RoboDK station: PickPlace_Delta_ABB.rdk

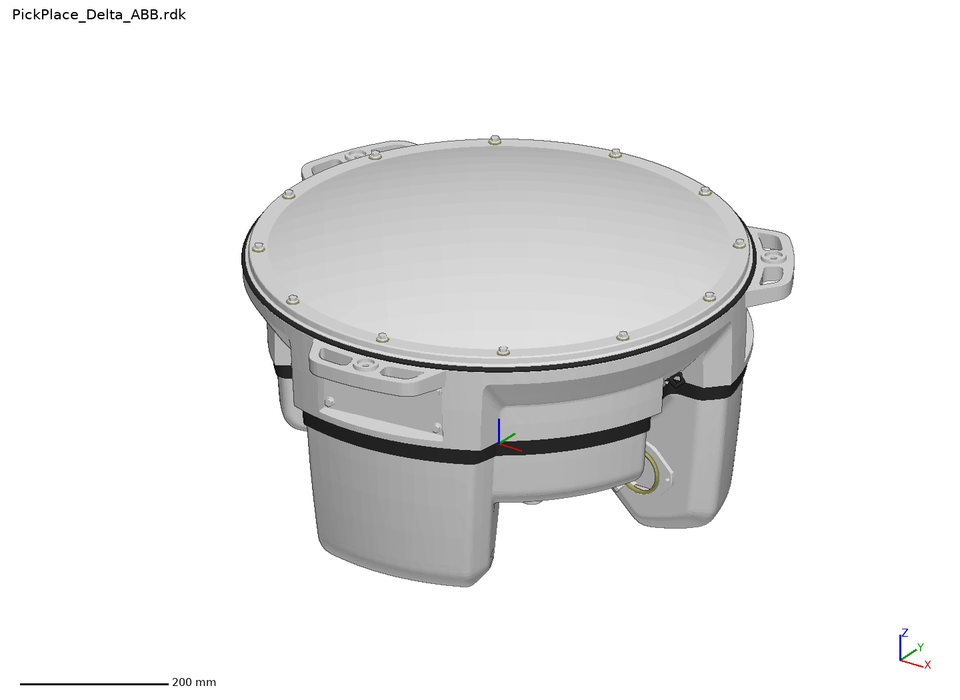
[picture v0: the station drawn from its stored meshes, robots at their saved joint values, targets as dots, program paths as lines]
Station PickPlace_Delta_ABB (saved by RoboDK 6.0.1). Poses are relative to the parent item; angles as X-Y-Z fixed-axis rotations.
Station parameters (name, value as stored): SICK WL4S Laser Sensor, 0, start_prox, 0
  - frame Conveyor Belt Wide (2m) Base at (0, 0, -10) mm
    - robot Conveyor Belt Wide (2m): 1 axes
        modified DH rows (alpha deg, a mm, theta deg, d mm): 0, 0, 0, 0 linear
        base shift (0, 0, 0) mm, rotated rx 0 ry 90 rz 0 deg
        joint limits [-900000] to [900000]; home [0]; saved at [-824508]
      - frame Conveyor Frame at (1954.3, 0, -10) mm
        - object Box at (897730.69, 156.17, 12.65) mm, rotated rx -0.59 ry -0.06 rz -23.58 deg, size 10 x 20 x 5 mm, geometry from box.sld
        - object Box at (897637.69, 177.81, 12.44) mm, rotated rx -0.3 ry 0.51 rz 41.51 deg, size 10 x 20 x 5 mm, geometry from box.sld
        - object Box at (897468.69, 142.01, 12.79) mm, rotated rx -0.52 ry 0.28 rz 10.42 deg, size 10 x 20 x 5 mm, geometry from box.sld
        - object Box at (897370.7, 94.71, 13.25) mm, rotated rx -0.59 ry 0.03 rz -15.02 deg, size 10 x 20 x 5 mm, geometry from box.sld
        - object Box at (897268.7, 59.56, 13.6) mm, rotated rx -0.59 ry -0.09 rz -26.61 deg, size 10 x 20 x 5 mm, geometry from box.sld
        - object Box at (897066.69, 179.61, 12.42) mm, rotated rx -0.4 ry 0.44 rz 29.48 deg, size 10 x 20 x 5 mm, geometry from box.sld
        - object Box at (896960.69, 179.12, 12.42) mm, rotated rx -0.29 ry 0.52 rz 42.93 deg, size 10 x 20 x 5 mm, geometry from box.sld
        - object Box at (896886.7, 104.97, 13.15) mm, rotated rx -0.55 ry 0.22 rz 3.61 deg, size 10 x 20 x 5 mm, geometry from box.sld
        - object Box at (896794.7, 36.7, 13.82) mm, rotated rx -0.43 ry 0.41 rz 25.81 deg, size 10 x 20 x 5 mm, geometry from box.sld
        - object Box at (896686.7, 102.36, 13.18) mm, rotated rx -0.56 ry -0.21 rz -38.82 deg, size 10 x 20 x 5 mm, geometry from box.sld
        - object Box at (896480.69, 181.98, 12.39) mm, rotated rx -0.53 ry -0.26 rz -44.04 deg, size 10 x 20 x 5 mm, geometry from box.sld
        - object Box at (896386.7, 69.3, 13.5) mm, rotated rx -0.54 ry -0.24 rz -42.5 deg, size 10 x 20 x 5 mm, geometry from box.sld
        - object Box at (896271.7, 21, 13.98) mm, rotated rx -0.57 ry -0.15 rz -32.81 deg, size 10 x 20 x 5 mm, geometry from box.sld
        - object Box at (896066.7, 121.17, 12.99) mm, rotated rx -0.58 ry 0.12 rz -6.35 deg, size 10 x 20 x 5 mm, geometry from box.sld
        - object Box at (895875.7, 101.57, 13.19) mm, rotated rx -0.59 ry -0.02 rz -20.07 deg, size 10 x 20 x 5 mm, geometry from box.sld
        - object Box at (895769.69, 140.05, 12.81) mm, rotated rx -0.59 ry 0.01 rz -17.18 deg, size 10 x 20 x 5 mm, geometry from box.sld
        - object Box at (895559.7, 47.66, 13.72) mm, rotated rx -0.46 ry 0.38 rz 21.06 deg, size 10 x 20 x 5 mm, geometry from box.sld
        - object Box at (895483.69, 179.87, 12.41) mm, rotated rx -0.56 ry 0.2 rz 1.63 deg, size 10 x 20 x 5 mm, geometry from box.sld
        - object Box at (895370.7, 123.7, 12.97) mm, rotated rx -0.59 ry 0.04 rz -14.74 deg, size 10 x 20 x 5 mm, geometry from box.sld
        - object Box at (895264.7, 131.8, 12.89) mm, rotated rx -0.58 ry -0.14 rz -31.52 deg, size 10 x 20 x 5 mm, geometry from box.sld
        - object Box at (895176.7, 127.41, 12.93) mm, rotated rx -0.59 ry -0.01 rz -19.42 deg, size 10 x 20 x 5 mm, geometry from box.sld
        - object Box at (895070.69, 148.83, 12.72) mm, rotated rx -0.59 ry 0.04 rz -13.82 deg, size 10 x 20 x 5 mm, geometry from box.sld
        - object Box at (894830.7, 134.47, 12.86) mm, rotated rx -0.55 ry -0.21 rz -39.3 deg, size 10 x 20 x 5 mm, geometry from box.sld
        - object Box at (894736.69, 145.17, 12.76) mm, rotated rx -0.58 ry 0.12 rz -6.93 deg, size 10 x 20 x 5 mm, geometry from box.sld
        - object Box at (894651.7, 66.02, 13.54) mm, rotated rx -0.57 ry -0.15 rz -32.83 deg, size 10 x 20 x 5 mm, geometry from box.sld
        - object Box at (894556.7, 45.28, 13.74) mm, rotated rx -0.42 ry 0.42 rz 26.95 deg, size 10 x 20 x 5 mm, geometry from box.sld
        - object Box at (894429.7, 71.11, 13.49) mm, rotated rx -0.56 ry -0.2 rz -37.64 deg, size 10 x 20 x 5 mm, geometry from box.sld
        - object Box at (894341.69, 182.71, 12.39) mm, rotated rx -0.59 ry 0.01 rz -17.44 deg, size 10 x 20 x 5 mm, geometry from box.sld
        - object Box at (894244.7, 91.87, 13.28) mm, rotated rx -0.54 ry -0.24 rz -42.33 deg, size 10 x 20 x 5 mm, geometry from box.sld
        - object Box at (893942.7, 111.28, 13.09) mm, rotated rx -0.52 ry 0.28 rz 9.97 deg, size 10 x 20 x 5 mm, geometry from box.sld
        - object Box at (893859.7, 78.43, 13.41) mm, rotated rx -0.59 ry 0.05 rz -12.95 deg, size 10 x 20 x 5 mm, geometry from box.sld
        - object Box at (893731.69, 182.25, 12.39) mm, rotated rx -0.59 ry -0.05 rz -23.07 deg, size 10 x 20 x 5 mm, geometry from box.sld
        - object Box at (893626.69, 198.26, 12.23) mm, rotated rx -0.44 ry 0.4 rz 24.46 deg, size 10 x 20 x 5 mm, geometry from box.sld
        - object Box at (893339.7, 130.91, 12.9) mm, rotated rx -0.43 ry 0.41 rz 25.41 deg, size 10 x 20 x 5 mm, geometry from box.sld
        - object Box at (893114.69, 144.51, 12.76) mm, rotated rx -0.59 ry -0.04 rz -22.45 deg, size 10 x 20 x 5 mm, geometry from box.sld
        - object Box at (893046.7, 53.65, 13.66) mm, rotated rx -0.57 ry 0.15 rz -3.55 deg, size 10 x 20 x 5 mm, geometry from box.sld
        - object Box at (892837.69, 193.79, 12.28) mm, rotated rx -0.41 ry 0.43 rz 28.71 deg, size 10 x 20 x 5 mm, geometry from box.sld
        - object Box at (892611.7, 108.11, 13.12) mm, rotated rx -0.42 ry 0.42 rz 26.96 deg, size 10 x 20 x 5 mm, geometry from box.sld
        - object Box at (892480.7, 68.86, 13.51) mm, rotated rx -0.51 ry 0.3 rz 12.73 deg, size 10 x 20 x 5 mm, geometry from box.sld
        - object Box at (892369.7, 112.85, 13.07) mm, rotated rx -0.59 ry 0.02 rz -16.52 deg, size 10 x 20 x 5 mm, geometry from box.sld
        - object Box at (892237.7, 18.64, 14) mm, rotated rx -0.59 ry 0.06 rz -11.95 deg, size 10 x 20 x 5 mm, geometry from box.sld
        - object Box at (892122.69, 158.92, 12.62) mm, rotated rx -0.43 ry 0.41 rz 25.04 deg, size 10 x 20 x 5 mm, geometry from box.sld
        - object Box at (892026.7, 94.47, 13.26) mm, rotated rx -0.59 ry 0.07 rz -11.43 deg, size 10 x 20 x 5 mm, geometry from box.sld
        - object Box at (891747.7, 66.89, 13.53) mm, rotated rx -0.59 ry -0.02 rz -20.16 deg, size 10 x 20 x 5 mm, geometry from box.sld
        - object Box at (891542.69, 140.71, 12.8) mm, rotated rx -0.42 ry 0.42 rz 26.92 deg, size 10 x 20 x 5 mm, geometry from box.sld
        - object Box at (891444.69, 197.73, 12.24) mm, rotated rx -0.3 ry 0.51 rz 41.43 deg, size 10 x 20 x 5 mm, geometry from box.sld
        - object Box at (891351.7, 42.87, 13.76) mm, rotated rx -0.54 ry -0.24 rz -41.92 deg, size 10 x 20 x 5 mm, geometry from box.sld
        - object Box at (891043.69, 177.02, 12.44) mm, rotated rx -0.57 ry -0.17 rz -35.25 deg, size 10 x 20 x 5 mm, geometry from box.sld
        - object Box at (890826.69, 146.16, 12.75) mm, rotated rx -0.57 ry -0.16 rz -33.48 deg, size 10 x 20 x 5 mm, geometry from box.sld
        - object Box at (890637.7, 55.66, 13.64) mm, rotated rx -0.58 ry -0.13 rz -30.72 deg, size 10 x 20 x 5 mm, geometry from box.sld
        - object Box at (890524.69, 170.49, 12.51) mm, rotated rx -0.57 ry -0.16 rz -33.37 deg, size 10 x 20 x 5 mm, geometry from box.sld
        - object Box at (890376.69, 167.1, 12.54) mm, rotated rx -0.58 ry -0.12 rz -30.29 deg, size 10 x 20 x 5 mm, geometry from box.sld
        - object Box at (890243.7, 28.37, 13.91) mm, rotated rx -0.59 ry -0.03 rz -21.44 deg, size 10 x 20 x 5 mm, geometry from box.sld
        - object Box at (890087.7, 32.55, 13.87) mm, rotated rx -0.58 ry -0.14 rz -31.77 deg, size 10 x 20 x 5 mm, geometry from box.sld
        - object Box at (889842.7, 52.41, 13.67) mm, rotated rx -0.49 ry 0.33 rz 15.68 deg, size 10 x 20 x 5 mm, geometry from box.sld
        - object Box at (889568.7, 81.43, 13.38) mm, rotated rx -0.43 ry 0.41 rz 25.3 deg, size 10 x 20 x 5 mm, geometry from box.sld
        - object Box at (889310.7, 27.98, 13.91) mm, rotated rx -0.57 ry 0.18 rz -0.36 deg, size 10 x 20 x 5 mm, geometry from box.sld
        - object Box at (889224.69, 159.39, 12.62) mm, rotated rx -0.5 ry 0.32 rz 14.94 deg, size 10 x 20 x 5 mm, geometry from box.sld
        - object Box at (888940.7, 109.26, 13.11) mm, rotated rx -0.58 ry 0.13 rz -5.05 deg, size 10 x 20 x 5 mm, geometry from box.sld
        - object Box at (888797.7, 63.43, 13.56) mm, rotated rx -0.32 ry 0.5 rz 38.96 deg, size 10 x 20 x 5 mm, geometry from box.sld
        - object Box at (888564.7, 67.11, 13.52) mm, rotated rx -0.39 ry 0.45 rz 31 deg, size 10 x 20 x 5 mm, geometry from box.sld
        - object Box at (888277.69, 157.91, 12.63) mm, rotated rx -0.51 ry 0.31 rz 12.91 deg, size 10 x 20 x 5 mm, geometry from box.sld
        - object Box at (888179.7, 88.13, 13.32) mm, rotated rx -0.53 ry 0.26 rz 8.19 deg, size 10 x 20 x 5 mm, geometry from box.sld
        - object Box at (888049.69, 160.71, 12.6) mm, rotated rx -0.59 ry -0.04 rz -22.46 deg, size 10 x 20 x 5 mm, geometry from box.sld
        - object Box at (887779.69, 175.73, 12.46) mm, rotated rx -0.56 ry 0.18 rz -0.25 deg, size 10 x 20 x 5 mm, geometry from box.sld
        - object Box at (887507.7, 34.78, 13.84) mm, rotated rx -0.55 ry 0.23 rz 5.02 deg, size 10 x 20 x 5 mm, geometry from box.sld
        - object Box at (887341.69, 183.19, 12.38) mm, rotated rx -0.35 ry 0.48 rz 36.16 deg, size 10 x 20 x 5 mm, geometry from box.sld
        - object Box at (887031.7, 18.9, 14) mm, rotated rx -0.59 ry -0.08 rz -26.28 deg, size 10 x 20 x 5 mm, geometry from box.sld
        - object Box at (886865.69, 175.99, 12.45) mm, rotated rx -0.58 ry 0.15 rz -3.88 deg, size 10 x 20 x 5 mm, geometry from box.sld
        - object Box at (886728.7, 132.72, 12.88) mm, rotated rx -0.47 ry 0.36 rz 18.81 deg, size 10 x 20 x 5 mm, geometry from box.sld
        - object Box at (886614.7, 70.74, 13.49) mm, rotated rx -0.56 ry 0.2 rz 1.77 deg, size 10 x 20 x 5 mm, geometry from box.sld
        - object Box at (886478.7, 44.32, 13.75) mm, rotated rx -0.58 ry -0.11 rz -29.31 deg, size 10 x 20 x 5 mm, geometry from box.sld
        - object Box at (886356.7, 71.95, 13.48) mm, rotated rx -0.51 ry 0.31 rz 13.14 deg, size 10 x 20 x 5 mm, geometry from box.sld
        - object Box at (886087.7, 108.74, 13.12) mm, rotated rx -0.58 ry -0.13 rz -31.01 deg, size 10 x 20 x 5 mm, geometry from box.sld
        - object Box at (885692.69, 167.79, 12.53) mm, rotated rx -0.59 ry -0.01 rz -18.94 deg, size 10 x 20 x 5 mm, geometry from box.sld
        - object Box at (885279.7, 93.51, 13.26) mm, rotated rx -0.57 ry -0.17 rz -35.18 deg, size 10 x 20 x 5 mm, geometry from box.sld
        - object Box at (885168.7, 33.77, 13.85) mm, rotated rx -0.59 ry 0.09 rz -9.53 deg, size 10 x 20 x 5 mm, geometry from box.sld
        - object Box at (884865.7, 95.2, 13.25) mm, rotated rx -0.59 ry -0.1 rz -27.76 deg, size 10 x 20 x 5 mm, geometry from box.sld
        - object Box at (884481.69, 195.64, 12.26) mm, rotated rx -0.59 ry 0.05 rz -13.6 deg, size 10 x 20 x 5 mm, geometry from box.sld
        - object Box at (884238.7, 13.58, 14.05) mm, rotated rx -0.29 ry 0.52 rz 42.46 deg, size 10 x 20 x 5 mm, geometry from box.sld
        - object Box at (883600.69, 168.73, 12.52) mm, rotated rx -0.39 ry 0.45 rz 31.19 deg, size 10 x 20 x 5 mm, geometry from box.sld
        - object Box at (883471.69, 175.1, 12.46) mm, rotated rx -0.56 ry -0.19 rz -36.67 deg, size 10 x 20 x 5 mm, geometry from box.sld
        - object Box at (883117.7, 8.08, 14.11) mm, rotated rx -0.59 ry 0 rz -18.33 deg, size 10 x 20 x 5 mm, geometry from box.sld
        - object Box at (882411.69, 148.37, 12.72) mm, rotated rx -0.37 ry 0.47 rz 33.68 deg, size 10 x 20 x 5 mm, geometry from box.sld
        - object Box at (881994.69, 149.13, 12.72) mm, rotated rx -0.55 ry -0.21 rz -39.37 deg, size 10 x 20 x 5 mm, geometry from box.sld
        - object Box at (881721.7, 36.8, 13.82) mm, rotated rx -0.56 ry -0.18 rz -36.26 deg, size 10 x 20 x 5 mm, geometry from box.sld
        - object Box at (881386.69, 181.59, 12.4) mm, rotated rx -0.48 ry 0.34 rz 17.23 deg, size 10 x 20 x 5 mm, geometry from box.sld
        - object Box at (881076.7, 104.94, 13.15) mm, rotated rx -0.58 ry 0.14 rz -4.54 deg, size 10 x 20 x 5 mm, geometry from box.sld
        - object Box at (880927.7, 105.79, 13.14) mm, rotated rx -0.59 ry -0.05 rz -23.21 deg, size 10 x 20 x 5 mm, geometry from box.sld
        - object Box at (880633.7, 82.69, 13.37) mm, rotated rx -0.58 ry 0.15 rz -3.91 deg, size 10 x 20 x 5 mm, geometry from box.sld
        - object Box at (880250.7, 100.17, 13.2) mm, rotated rx -0.35 ry 0.48 rz 36.02 deg, size 10 x 20 x 5 mm, geometry from box.sld
        - object Box at (879967.7, 8.92, 14.1) mm, rotated rx -0.34 ry 0.49 rz 36.88 deg, size 10 x 20 x 5 mm, geometry from box.sld
        - object Box at (879702.69, 197.41, 12.24) mm, rotated rx -0.54 ry 0.24 rz 5.94 deg, size 10 x 20 x 5 mm, geometry from box.sld
        - object Box at (879327.7, 134.52, 12.86) mm, rotated rx -0.31 ry 0.51 rz 40.25 deg, size 10 x 20 x 5 mm, geometry from box.sld
        - object Box at (879021.7, 66.06, 13.54) mm, rotated rx -0.59 ry -0.09 rz -26.74 deg, size 10 x 20 x 5 mm, geometry from box.sld
        - object Box at (878707.7, 123.22, 12.97) mm, rotated rx -0.3 ry 0.51 rz 41.76 deg, size 10 x 20 x 5 mm, geometry from box.sld
        - object Box at (878458.7, 26.6, 13.92) mm, rotated rx -0.38 ry 0.46 rz 32.24 deg, size 10 x 20 x 5 mm, geometry from box.sld
        - object Box at (878137.69, 148.25, 12.73) mm, rotated rx -0.36 ry 0.47 rz 34.26 deg, size 10 x 20 x 5 mm, geometry from box.sld
        - object Box at (877571.7, 84.32, 13.36) mm, rotated rx -0.33 ry 0.5 rz 38.45 deg, size 10 x 20 x 5 mm, geometry from box.sld
        - object Box at (877259.69, 194, 12.28) mm, rotated rx -0.49 ry 0.33 rz 15.69 deg, size 10 x 20 x 5 mm, geometry from box.sld
        - object Box at (877049.69, 140.02, 12.81) mm, rotated rx -0.59 ry 0.01 rz -17.21 deg, size 10 x 20 x 5 mm, geometry from box.sld
        - object Box at (876618.69, 160.9, 12.6) mm, rotated rx -0.56 ry -0.21 rz -38.5 deg, size 10 x 20 x 5 mm, geometry from box.sld
        - object Box at (876232.69, 160.62, 12.6) mm, rotated rx -0.52 ry 0.28 rz 10.27 deg, size 10 x 20 x 5 mm, geometry from box.sld
        - object Box at (876057.7, 87.66, 13.32) mm, rotated rx -0.56 ry -0.21 rz -38.4 deg, size 10 x 20 x 5 mm, geometry from box.sld
        - object Box at (875735.69, 153.67, 12.67) mm, rotated rx -0.57 ry 0.17 rz -1.28 deg, size 10 x 20 x 5 mm, geometry from box.sld
        - object Box at (875385.7, 12.69, 14.06) mm, rotated rx -0.52 ry 0.29 rz 10.64 deg, size 10 x 20 x 5 mm, geometry from box.sld
        - object Box at (874877.7, 46, 13.73) mm, rotated rx -0.46 ry 0.37 rz 20.28 deg, size 10 x 20 x 5 mm, geometry from box.sld
        - object Box at (874555.69, 151.65, 12.69) mm, rotated rx -0.58 ry -0.14 rz -31.99 deg, size 10 x 20 x 5 mm, geometry from box.sld
        - object Box at (873807.69, 173.16, 12.48) mm, rotated rx -0.28 ry 0.52 rz 43.49 deg, size 10 x 20 x 5 mm, geometry from box.sld
        - object Box at (872936.7, 49.92, 13.69) mm, rotated rx -0.34 ry 0.49 rz 36.91 deg, size 10 x 20 x 5 mm, geometry from box.sld
        - object Box at (872785.69, 161.75, 12.59) mm, rotated rx -0.59 ry 0.09 rz -9.24 deg, size 10 x 20 x 5 mm, geometry from box.sld
        - object Box at (872664.7, 91.07, 13.29) mm, rotated rx -0.52 ry 0.29 rz 11.2 deg, size 10 x 20 x 5 mm, geometry from box.sld
        - object Box at (872500.7, 40.63, 13.79) mm, rotated rx -0.59 ry 0.06 rz -12.41 deg, size 10 x 20 x 5 mm, geometry from box.sld
        - object Box at (872142.7, 105.29, 13.15) mm, rotated rx -0.5 ry 0.32 rz 14.54 deg, size 10 x 20 x 5 mm, geometry from box.sld
        - object Box at (871888.7, 15.8, 14.03) mm, rotated rx -0.53 ry -0.27 rz -44.74 deg, size 10 x 20 x 5 mm, geometry from box.sld
        - object Box at (871587.7, 7.86, 14.11) mm, rotated rx -0.51 ry 0.3 rz 12.38 deg, size 10 x 20 x 5 mm, geometry from box.sld
        - object Box at (870973.69, 136.14, 12.85) mm, rotated rx -0.42 ry 0.42 rz 26.47 deg, size 10 x 20 x 5 mm, geometry from box.sld
        - object Box at (869775.7, 70.75, 13.49) mm, rotated rx -0.38 ry 0.46 rz 32.57 deg, size 10 x 20 x 5 mm, geometry from box.sld
        - object Box at (869038.69, 182.24, 12.39) mm, rotated rx -0.55 ry -0.21 rz -39.23 deg, size 10 x 20 x 5 mm, geometry from box.sld
        - object Box at (868878.7, 50.82, 13.69) mm, rotated rx -0.59 ry 0.03 rz -15.61 deg, size 10 x 20 x 5 mm, geometry from box.sld
        - object Box at (868388.7, 14.54, 14.04) mm, rotated rx -0.57 ry 0.15 rz -3.36 deg, size 10 x 20 x 5 mm, geometry from box.sld
        - object Box at (867960.7, 83.04, 13.37) mm, rotated rx -0.52 ry 0.28 rz 9.96 deg, size 10 x 20 x 5 mm, geometry from box.sld
        - object Box at (867636.7, 10.32, 14.08) mm, rotated rx -0.4 ry 0.44 rz 29.65 deg, size 10 x 20 x 5 mm, geometry from box.sld
        - object Box at (867059.69, 162.68, 12.58) mm, rotated rx -0.58 ry -0.11 rz -28.52 deg, size 10 x 20 x 5 mm, geometry from box.sld
        - object Box at (866931.7, 128.82, 12.92) mm, rotated rx -0.55 ry 0.21 rz 2.62 deg, size 10 x 20 x 5 mm, geometry from box.sld
        - object Box at (866587.69, 156.78, 12.64) mm, rotated rx -0.47 ry 0.36 rz 19.55 deg, size 10 x 20 x 5 mm, geometry from box.sld
        - object Box at (866076.69, 184.18, 12.37) mm, rotated rx -0.59 ry 0.04 rz -14.44 deg, size 10 x 20 x 5 mm, geometry from box.sld
        - object Box at (865379.7, 5.34, 14.13) mm, rotated rx -0.58 ry -0.13 rz -30.77 deg, size 10 x 20 x 5 mm, geometry from box.sld
        - object Box at (865212.69, 149.76, 12.71) mm, rotated rx -0.56 ry -0.2 rz -38.32 deg, size 10 x 20 x 5 mm, geometry from box.sld
        - object Box at (864790.7, 7.34, 14.11) mm, rotated rx -0.59 ry 0.07 rz -11.85 deg, size 10 x 20 x 5 mm, geometry from box.sld
        - object Box at (864117.7, 14.14, 14.05) mm, rotated rx -0.4 ry 0.44 rz 29.12 deg, size 10 x 20 x 5 mm, geometry from box.sld
        - object Box at (864010.69, 143.76, 12.77) mm, rotated rx -0.59 ry 0 rz -18.52 deg, size 10 x 20 x 5 mm, geometry from box.sld
        - object Box at (863847.69, 186.35, 12.35) mm, rotated rx -0.54 ry -0.24 rz -42.33 deg, size 10 x 20 x 5 mm, geometry from box.sld
        - object Box at (863773.7, 56.85, 13.63) mm, rotated rx -0.53 ry -0.27 rz -44.81 deg, size 10 x 20 x 5 mm, geometry from box.sld
        - object Box at (863691.7, 42.47, 13.77) mm, rotated rx -0.57 ry -0.16 rz -34.11 deg, size 10 x 20 x 5 mm, geometry from box.sld
        - object Box at (863609.7, 44.95, 13.74) mm, rotated rx -0.5 ry 0.33 rz 15.05 deg, size 10 x 20 x 5 mm, geometry from box.sld
        - object Box at (863543.7, 34.25, 13.85) mm, rotated rx -0.51 ry 0.31 rz 13.03 deg, size 10 x 20 x 5 mm, geometry from box.sld
        - object Box at (863468.7, 76.02, 13.44) mm, rotated rx -0.59 ry 0.1 rz -8.77 deg, size 10 x 20 x 5 mm, geometry from box.sld
        - object Box at (863299.7, 107.42, 13.13) mm, rotated rx -0.55 ry -0.21 rz -39.28 deg, size 10 x 20 x 5 mm, geometry from box.sld
        - object Box at (863239.69, 195.88, 12.26) mm, rotated rx -0.29 ry 0.52 rz 42.8 deg, size 10 x 20 x 5 mm, geometry from box.sld
        - object Box at (863168.7, 58.58, 13.61) mm, rotated rx -0.58 ry 0.15 rz -3.89 deg, size 10 x 20 x 5 mm, geometry from box.sld
        - object Box at (863074.69, 157.27, 12.64) mm, rotated rx -0.57 ry 0.17 rz -1.09 deg, size 10 x 20 x 5 mm, geometry from box.sld
        - object Box at (862995.7, 21.42, 13.97) mm, rotated rx -0.59 ry 0.1 rz -8.62 deg, size 10 x 20 x 5 mm, geometry from box.sld
        - object Box at (862844.69, 190.46, 12.31) mm, rotated rx -0.47 ry 0.37 rz 19.8 deg, size 10 x 20 x 5 mm, geometry from box.sld
        - object Box at (862697.7, 12.52, 14.06) mm, rotated rx -0.55 ry 0.22 rz 3.49 deg, size 10 x 20 x 5 mm, geometry from box.sld
        - object Box at (862605.7, 93.15, 13.27) mm, rotated rx -0.43 ry 0.41 rz 25.14 deg, size 10 x 20 x 5 mm, geometry from box.sld
        - object Box at (862511.69, 173.93, 12.47) mm, rotated rx -0.49 ry 0.33 rz 15.38 deg, size 10 x 20 x 5 mm, geometry from box.sld
        - object Box at (862445.69, 170.13, 12.51) mm, rotated rx -0.56 ry -0.21 rz -38.76 deg, size 10 x 20 x 5 mm, geometry from box.sld
        - object Box at (862285.69, 194.2, 12.27) mm, rotated rx -0.59 ry -0.02 rz -20.35 deg, size 10 x 20 x 5 mm, geometry from box.sld
        - object Box at (862212.7, 48.11, 13.71) mm, rotated rx -0.53 ry 0.26 rz 8.23 deg, size 10 x 20 x 5 mm, geometry from box.sld
        - object Box at (862077.7, 40.74, 13.78) mm, rotated rx -0.57 ry -0.15 rz -33.02 deg, size 10 x 20 x 5 mm, geometry from box.sld
        - object Box at (862001.69, 144.78, 12.76) mm, rotated rx -0.59 ry -0.04 rz -21.98 deg, size 10 x 20 x 5 mm, geometry from box.sld
        - object Box at (861912.7, 129.98, 12.91) mm, rotated rx -0.41 ry 0.43 rz 27.6 deg, size 10 x 20 x 5 mm, geometry from box.sld
        - object Box at (861831.7, 111.46, 13.09) mm, rotated rx -0.56 ry -0.2 rz -37.82 deg, size 10 x 20 x 5 mm, geometry from box.sld
        - object Box at (861677.7, 88.75, 13.31) mm, rotated rx -0.59 ry 0.05 rz -13.53 deg, size 10 x 20 x 5 mm, geometry from box.sld
        - object Box at (861612.69, 197.69, 12.24) mm, rotated rx -0.59 ry -0.05 rz -22.69 deg, size 10 x 20 x 5 mm, geometry from box.sld
        - object Box at (861533.7, 55.71, 13.64) mm, rotated rx -0.59 ry 0.08 rz -10.75 deg, size 10 x 20 x 5 mm, geometry from box.sld
        - object Box at (861367.7, 89.81, 13.3) mm, rotated rx -0.46 ry 0.37 rz 20.67 deg, size 10 x 20 x 5 mm, geometry from box.sld
        - object Box at (861299.7, 23.97, 13.95) mm, rotated rx -0.59 ry 0.05 rz -12.94 deg, size 10 x 20 x 5 mm, geometry from box.sld
        - object Box at (861219.7, 9.88, 14.09) mm, rotated rx -0.53 ry 0.26 rz 7.95 deg, size 10 x 20 x 5 mm, geometry from box.sld
        - object Box at (861142.7, 51.83, 13.68) mm, rotated rx -0.42 ry 0.42 rz 27.28 deg, size 10 x 20 x 5 mm, geometry from box.sld
        - object Box at (861076.7, 108.48, 13.12) mm, rotated rx -0.55 ry -0.21 rz -38.97 deg, size 10 x 20 x 5 mm, geometry from box.sld
        - object Box at (860992.69, 187.44, 12.34) mm, rotated rx -0.59 ry -0.04 rz -22.25 deg, size 10 x 20 x 5 mm, geometry from box.sld
        - object Box at (860907.7, 101.41, 13.19) mm, rotated rx -0.38 ry 0.46 rz 32.23 deg, size 10 x 20 x 5 mm, geometry from box.sld
        - object Box at (860818.7, 75.58, 13.44) mm, rotated rx -0.48 ry 0.35 rz 18.56 deg, size 10 x 20 x 5 mm, geometry from box.sld
        - object Box at (860742.7, 42.49, 13.77) mm, rotated rx -0.47 ry 0.37 rz 20.23 deg, size 10 x 20 x 5 mm, geometry from box.sld
        - object Box at (860572.7, 93.25, 13.27) mm, rotated rx -0.28 ry 0.52 rz 43.65 deg, size 10 x 20 x 5 mm, geometry from box.sld
        - object Box at (860493.7, 47.45, 13.72) mm, rotated rx -0.56 ry 0.2 rz 1.93 deg, size 10 x 20 x 5 mm, geometry from box.sld
        - object Box at (860416.7, 72.1, 13.48) mm, rotated rx -0.56 ry -0.2 rz -37.75 deg, size 10 x 20 x 5 mm, geometry from box.sld
        - object Box at (860244.69, 202.97, 12.19) mm, rotated rx -0.58 ry -0.12 rz -30.25 deg, size 10 x 20 x 5 mm, geometry from box.sld
        - object Box at (860096.7, 47.66, 13.72) mm, rotated rx -0.59 ry -0.04 rz -22.39 deg, size 10 x 20 x 5 mm, geometry from box.sld
        - object Box at (860019.7, 98.6, 13.21) mm, rotated rx -0.45 ry 0.39 rz 23.07 deg, size 10 x 20 x 5 mm, geometry from box.sld
        - object Box at (859926.7, 66.26, 13.53) mm, rotated rx -0.54 ry -0.24 rz -42.09 deg, size 10 x 20 x 5 mm, geometry from box.sld
        - object Box at (859832.69, 186.44, 12.35) mm, rotated rx -0.55 ry -0.23 rz -41.1 deg, size 10 x 20 x 5 mm, geometry from box.sld
        - object Box at (859742.69, 188.27, 12.33) mm, rotated rx -0.34 ry 0.49 rz 36.82 deg, size 10 x 20 x 5 mm, geometry from box.sld
        - object Box at (859608.7, 60.54, 13.59) mm, rotated rx -0.44 ry 0.39 rz 23.51 deg, size 10 x 20 x 5 mm, geometry from box.sld
        - object Box at (859505.7, 104.17, 13.16) mm, rotated rx -0.59 ry 0.1 rz -8.48 deg, size 10 x 20 x 5 mm, geometry from box.sld
        - object Box at (859448.7, 129.15, 12.91) mm, rotated rx -0.53 ry -0.27 rz -44.76 deg, size 10 x 20 x 5 mm, geometry from box.sld
        - object Box at (859363.7, 97.67, 13.22) mm, rotated rx -0.57 ry -0.15 rz -33.2 deg, size 10 x 20 x 5 mm, geometry from box.sld
        - object Box at (859297.7, 133.43, 12.87) mm, rotated rx -0.59 ry -0.1 rz -27.76 deg, size 10 x 20 x 5 mm, geometry from box.sld
        - object Box at (859222.69, 179.69, 12.42) mm, rotated rx -0.55 ry -0.22 rz -39.91 deg, size 10 x 20 x 5 mm, geometry from box.sld
        - object Box at (859139.7, 100.3, 13.2) mm, rotated rx -0.58 ry 0.1 rz -8 deg, size 10 x 20 x 5 mm, geometry from box.sld
        - object Box at (858984.7, 92.61, 13.27) mm, rotated rx -0.32 ry 0.5 rz 39.39 deg, size 10 x 20 x 5 mm, geometry from box.sld
        - object Box at (858921.7, 78.7, 13.41) mm, rotated rx -0.38 ry 0.46 rz 32.5 deg, size 10 x 20 x 5 mm, geometry from box.sld
        - object Box at (858838.69, 182.91, 12.38) mm, rotated rx -0.42 ry 0.42 rz 27.15 deg, size 10 x 20 x 5 mm, geometry from box.sld
        - object Box at (858747.7, 41.89, 13.77) mm, rotated rx -0.59 ry -0.1 rz -27.61 deg, size 10 x 20 x 5 mm, geometry from box.sld
        - object Box at (858681.7, 26.61, 13.92) mm, rotated rx -0.55 ry -0.22 rz -39.6 deg, size 10 x 20 x 5 mm, geometry from box.sld
        - object Box at (858608.7, 106.46, 13.14) mm, rotated rx -0.59 ry -0.02 rz -19.7 deg, size 10 x 20 x 5 mm, geometry from box.sld
        - object Box at (858527.7, 43.27, 13.76) mm, rotated rx -0.55 ry -0.22 rz -40.16 deg, size 10 x 20 x 5 mm, geometry from box.sld
        - object Box at (858436.69, 147.53, 12.73) mm, rotated rx -0.38 ry 0.46 rz 32.63 deg, size 10 x 20 x 5 mm, geometry from box.sld
        - object Box at (858338.7, 95.37, 13.25) mm, rotated rx -0.46 ry 0.38 rz 21.04 deg, size 10 x 20 x 5 mm, geometry from box.sld
        - object Box at (858264.7, 16.13, 14.03) mm, rotated rx -0.34 ry 0.49 rz 37.01 deg, size 10 x 20 x 5 mm, geometry from box.sld
        - object Box at (858197.69, 138.48, 12.82) mm, rotated rx -0.5 ry 0.33 rz 15.3 deg, size 10 x 20 x 5 mm, geometry from box.sld
        - object Box at (858126.69, 164.96, 12.56) mm, rotated rx -0.59 ry 0.05 rz -13.57 deg, size 10 x 20 x 5 mm, geometry from box.sld
        - object Box at (858041.7, 93.37, 13.27) mm, rotated rx -0.54 ry -0.25 rz -42.69 deg, size 10 x 20 x 5 mm, geometry from box.sld
        - object Box at (857953.7, 107.45, 13.13) mm, rotated rx -0.42 ry 0.42 rz 27.28 deg, size 10 x 20 x 5 mm, geometry from box.sld
        - object Box at (857885.7, 120.25, 13) mm, rotated rx -0.49 ry 0.34 rz 16.8 deg, size 10 x 20 x 5 mm, geometry from box.sld
        - object Box at (857816.7, 44.03, 13.75) mm, rotated rx -0.55 ry -0.21 rz -39.24 deg, size 10 x 20 x 5 mm, geometry from box.sld
        - object Box at (857717.7, 12.89, 14.06) mm, rotated rx -0.59 ry 0.04 rz -14.42 deg, size 10 x 20 x 5 mm, geometry from box.sld
        - object Box at (857640.7, 89.25, 13.31) mm, rotated rx -0.53 ry 0.28 rz 9.63 deg, size 10 x 20 x 5 mm, geometry from box.sld
        - object Box at (857557.69, 134.96, 12.86) mm, rotated rx -0.46 ry 0.38 rz 21.35 deg, size 10 x 20 x 5 mm, geometry from box.sld
        - object Box at (857493.69, 197, 12.25) mm, rotated rx -0.59 ry -0.04 rz -22.07 deg, size 10 x 20 x 5 mm, geometry from box.sld
        - object Box at (857413.7, 74.98, 13.45) mm, rotated rx -0.53 ry 0.26 rz 7.8 deg, size 10 x 20 x 5 mm, geometry from box.sld
        - object Box at (857347.69, 145.19, 12.76) mm, rotated rx -0.59 ry 0.08 rz -10.75 deg, size 10 x 20 x 5 mm, geometry from box.sld
        - object Box at (857259.7, 112.65, 13.08) mm, rotated rx -0.51 ry 0.3 rz 11.87 deg, size 10 x 20 x 5 mm, geometry from box.sld
        - object Box at (857189.7, 106.79, 13.13) mm, rotated rx -0.5 ry 0.32 rz 14.38 deg, size 10 x 20 x 5 mm, geometry from box.sld
        - object Box at (857120.7, 96.6, 13.23) mm, rotated rx -0.59 ry -0.08 rz -26.03 deg, size 10 x 20 x 5 mm, geometry from box.sld
        - object Box at (857045.7, 85.92, 13.34) mm, rotated rx -0.58 ry 0.14 rz -4.09 deg, size 10 x 20 x 5 mm, geometry from box.sld
        - object Box at (856958.7, 103.33, 13.17) mm, rotated rx -0.57 ry 0.15 rz -3.36 deg, size 10 x 20 x 5 mm, geometry from box.sld
        - object Box at (856875.69, 160.95, 12.6) mm, rotated rx -0.52 ry 0.29 rz 11.23 deg, size 10 x 20 x 5 mm, geometry from box.sld
    - frame Reference Box Frame at (60, 290, 366.5) mm
      - object ref_obj at (0, 0, 0) mm, size 252 x 305.4 x 216.7 mm, geometry from Box-12x10in-Closed.sld
      - object ref_lid at (-60, -186.65, 3.17) mm, rotated rx -0.56 ry 0.19 rz 0 deg, size 10 x 20 x 5 mm, geometry from box.sld
      - object ref_lid1 at (-60, -86.65, 3.17) mm, rotated rx -0.56 ry 0.19 rz 0 deg, size 10 x 20 x 5 mm, geometry from box.sld
    - object SICK WL4S Laser Sensor at (1954, -20, 370) mm, rotated rx 180 ry 0 rz 90 deg, size 683.3 x 45.2 x 12.5 mm, geometry from SICK-WL4S-Laser-Sensor.sld
    - object start_prox at (0, -20, 370) mm, rotated rx 180 ry 0 rz 90 deg, size 683.3 x 45.2 x 12.5 mm, geometry from SICK-WL4S-Laser-Sensor.sld
  - program MainProgram (5 instructions, listed below)
  - notes Description: <!DOCTYPE HTML PUBLIC "-//W3C//DTD HTML 4.0//EN" "http://www.w3.org/TR/REC-html40/strict.dtd">
<html><head><meta name="qrichtext" content="1" /><style type="text/css">
p, li { white-space: pre-wrap; }
</style></head><body style=" font-family:'MS Shell Dlg 2'; font-size:8.25pt; font-weight:400; font-style:normal;">
<p style=" margin-top:0px; margin-bottom:0px; margin-left:0px; margin-right:0px; -qt-block-indent:0; text-indent:0px;">This example demonstrates a conveyor simulation in RoboDK using Python scripting. A script generates boxes of varying sizes and positions while the conveyor moves continuously. A sensor detects when a box reaches the conveyor’s edge and stops the conveyor. The station showcases how conveyors, part generation, and sensor-based control can be simulated with the API.</p></body></html>
  - frame ABB IRB 360-1/800 4D Base at (1954.3, 143.51, 1521.09) mm
    - robot ABB IRB 360-1/800 4D: 4 axes, payload 1 kg, reach 400 mm, repeatability 0.04 mm, weight 120 kg
        joint limits [-42, -42, -42, -36000] to [99.5, 99.5, 99.5, 36000]; home [0, 0, 0, 0]; saved at [15.4, 15.4, 15.4, 0]
      - tool Tool 1, TCP at (0, 0, 0) mm
  - frame CamFrame at (1207.08, 136.9, 843.5) mm, rotated rx -180 ry -0.2 rz -0.44 deg
    - camera Camera 1
  - frame Frame 6 at (1375.31, 171.47, 367.78) mm
  - frame Frame 7 at (1050, 111.47, 400) mm
  - frame delete_box_frame at (2400, 111.47, 400) mm

--- program MainProgram (robot Conveyor Belt Wide (2m)) ---
  Call ConveyorReset
  Run SensorReader
  Set speed (25.0 mm/s)
  Run ConveyorRunner
  Run BoxSpawner
